(* IEC 61131-3 sources: volt/packages/volt-lsp-iec/test-corpus/lenze-mid/Device/Plc Logic/Application/Library Manager/CAA RTCLK, 21 files *)

(* ---- ERROR.dut ---- *)
TYPE ERROR :
(
	NO_ERROR := 0,
	FIRST_ERROR := 5700,
	TIME_OUT := 5701,
	NOT_AVAILABLE := 5702,
	TIME_NOT_VALID := 5703,
	WRONG_PARAMETER := 5704,
	ERROR_UNKNOWN := 5705,
	NOT_IMPLEMENTED := 5706,
	FIRST_MF := 5725,
	LAST_ERROR := 5749
);
END_TYPE

(* ---- PERIODE.dut ---- *)
TYPE PERIODE :
(
	UNKNOWN := 0,
	STANDARD := 1,
	DAYLIGHT := 2
);
END_TYPE

(* ---- PERIODE_INFO.dut ---- *)
TYPE PERIODE_INFO : RTCLK_PERIODE_INFO;
END_TYPE

(* ---- RTCLK_GETDATEANDTIME_PARAMS.dut ---- *)
TYPE RTCLK_GETDATEANDTIME_PARAMS :
STRUCT
	DTDATEANDTIME : DATE_AND_TIME;
	ETIMEZONE : PERIODE;
END_STRUCT
END_TYPE

(* ---- RTCLK_GETTIMEZONEINFORMATION_PARAMS.dut ---- *)
TYPE RTCLK_GETTIMEZONEINFORMATION_PARAMS :
STRUCT
	TZITIMEZONE : RTCLK_TIME_ZONE_INFO;
END_STRUCT
END_TYPE

(* ---- RTCLK_PERIODE_INFO.dut ---- *)
TYPE RTCLK_PERIODE_INFO :
STRUCT
	SNAME : STRING(32);
	TMDATE : RTCLK_SYSTEMTIME;
	IBIAS : INT;
END_STRUCT
END_TYPE

(* ---- RTCLK_SETDATEANDTIME_PARAMS.dut ---- *)
TYPE RTCLK_SETDATEANDTIME_PARAMS :
STRUCT
	DTDATEANDTIME : DATE_AND_TIME;
END_STRUCT
END_TYPE

(* ---- RTCLK_SETTIMEZONEINFORMATION_PARAMS.dut ---- *)
TYPE RTCLK_SETTIMEZONEINFORMATION_PARAMS :
STRUCT
	TZITIMEZONE : RTCLK_TIME_ZONE_INFO;
END_STRUCT
END_TYPE

(* ---- RTCLK_SYSTEMTIME.dut ---- *)
TYPE RTCLK_SYSTEMTIME :
STRUCT
	UIYEAR : UINT;
	UIMONTH : UINT;
	EWEEKDAY : WEEKDAY;
	UIDAY : UINT;
	UIHOUR : UINT;
	UIMINUTE : UINT;
	UISECOND : UINT;
END_STRUCT
END_TYPE

(* ---- RTCLK_TIME_ZONE_INFO.dut ---- *)
TYPE RTCLK_TIME_ZONE_INFO :
STRUCT
	IBIAS : INT;
	SPERIODE : ARRAY [1..2] OF RTCLK_PERIODE_INFO;
END_STRUCT
END_TYPE

(* ---- SYSTEMTIME.dut ---- *)
TYPE SYSTEMTIME : RTCLK_SYSTEMTIME;
END_TYPE

(* ---- TIME_ZONE_INFO.dut ---- *)
TYPE TIME_ZONE_INFO : RTCLK_TIME_ZONE_INFO;
END_TYPE

(* ---- WEEKDAY.dut ---- *)
TYPE WEEKDAY :
(
	SUNDAY := 0,
	MONDAY := 1,
	TUESDAY := 2,
	WEDNESDAY := 3,
	THURSDAY := 4,
	FRIDAY := 5,
	SATURDAY := 6
);
END_TYPE

(* ---- PROPERTYCONSTANTS.gvl ---- *)
VAR_GLOBAL
	GC_WTIMEZONESUPPORT : WORD := 1;
END_VAR

(* ---- VERSIONCONSTANTS.gvl ---- *)
VAR_GLOBAL
	GC_BYVERSION : BYTE := 1;
	GC_BYVERSION_1 : BYTE := 0;
END_VAR

(* ---- GETPROPERTY.pou ---- *)
FUNCTION GETPROPERTY : __XWORD
VAR_INPUT
	WPROPERTY : WORD;
END_VAR
END_FUNCTION

(* ---- GETSUPPLIERVERSION.pou ---- *)
FUNCTION GETSUPPLIERVERSION : WORD
VAR_INPUT
	XDUMMY : BOOL;
END_VAR
END_FUNCTION

(* ---- GETDATEANDTIME.pou ---- *)
FUNCTION_BLOCK GETDATEANDTIME
VAR_INPUT
	XEXECUTE : BOOL;
END_VAR
VAR_OUTPUT
	XDONE : BOOL;
	XBUSY : BOOL;
	XERROR : BOOL;
	EERROR : ERROR;
	DTDATEANDTIME : DATE_AND_TIME;
	ETIMEZONE : PERIODE;
END_VAR
VAR
	XPREVIOUSEXECUTE : BOOL;
	XPREVIOUSABORTINPROGRESS : BOOL;
	XABORTINPROGRESS : BOOL;
	IERROR : INT;
	HJOB : CAA.HANDLE;
	PGETDATEANDTIMEPARAMS : POINTER TO RTCLK_GETDATEANDTIME_PARAMS;
	STATEJOB : ASM.STATE;
	DWETRIGCLASS : __XWORD;
END_VAR
END_FUNCTION_BLOCK

METHOD FB_EXIT : BOOL
VAR_INPUT
	BINCOPYCODE : BOOL;
END_VAR
END_METHOD

METHOD FB_INIT : BOOL
VAR_INPUT
	BINITRETAINS : BOOL;
	BINCOPYCODE : BOOL;
END_VAR
END_METHOD

(* ---- GETTIMEZONEINFORMATION.pou ---- *)
FUNCTION_BLOCK GETTIMEZONEINFORMATION
VAR_INPUT
	XEXECUTE : BOOL;
END_VAR
VAR_OUTPUT
	XDONE : BOOL;
	XBUSY : BOOL;
	XERROR : BOOL;
	EERROR : ERROR;
	TZIINFO : RTCLK_TIME_ZONE_INFO;
END_VAR
VAR
	XPREVIOUSEXECUTE : BOOL;
	XPREVIOUSABORTINPROGRESS : BOOL;
	XABORTINPROGRESS : BOOL;
	IERROR : INT;
	HJOB : CAA.HANDLE;
	PGETTIMEZONEINFORMATIONPARAMS : POINTER TO RTCLK_GETTIMEZONEINFORMATION_PARAMS;
	STATEJOB : ASM.STATE;
	DWETRIGCLASS : __XWORD;
END_VAR
END_FUNCTION_BLOCK

METHOD FB_EXIT : BOOL
VAR_INPUT
	BINCOPYCODE : BOOL;
END_VAR
END_METHOD

METHOD FB_INIT : BOOL
VAR_INPUT
	BINITRETAINS : BOOL;
	BINCOPYCODE : BOOL;
END_VAR
END_METHOD

(* ---- SETDATEANDTIME.pou ---- *)
FUNCTION_BLOCK SETDATEANDTIME
VAR_INPUT
	XEXECUTE : BOOL;
	DTDATEANDTIME : DATE_AND_TIME;
END_VAR
VAR_OUTPUT
	XDONE : BOOL;
	XBUSY : BOOL;
	XERROR : BOOL;
	EERROR : ERROR;
END_VAR
VAR
	XPREVIOUSEXECUTE : BOOL;
	XPREVIOUSABORTINPROGRESS : BOOL;
	XABORTINPROGRESS : BOOL;
	IERROR : INT;
	HJOB : CAA.HANDLE;
	PSETDATEANDTIMEPARAMS : POINTER TO RTCLK_SETDATEANDTIME_PARAMS;
	STATEJOB : ASM.STATE;
	DWETRIGCLASS : __XWORD;
END_VAR
END_FUNCTION_BLOCK

METHOD FB_EXIT : BOOL
VAR_INPUT
	BINCOPYCODE : BOOL;
END_VAR
END_METHOD

METHOD FB_INIT : BOOL
VAR_INPUT
	BINITRETAINS : BOOL;
	BINCOPYCODE : BOOL;
END_VAR
END_METHOD

(* ---- SETTIMEZONEINFORMATION.pou ---- *)
FUNCTION_BLOCK SETTIMEZONEINFORMATION
VAR_INPUT
	XEXECUTE : BOOL;
	TZIINFO : RTCLK_TIME_ZONE_INFO;
END_VAR
VAR_OUTPUT
	XDONE : BOOL;
	XBUSY : BOOL;
	XERROR : BOOL;
	EERROR : ERROR;
END_VAR
VAR
	XPREVIOUSEXECUTE : BOOL;
	XPREVIOUSABORTINPROGRESS : BOOL;
	XABORTINPROGRESS : BOOL;
	IERROR : INT;
	HJOB : CAA.HANDLE;
	PSETTIMEZONEINFORMATIONPARAMS : POINTER TO RTCLK_SETTIMEZONEINFORMATION_PARAMS;
	STATEJOB : ASM.STATE;
	DWETRIGCLASS : __XWORD;
END_VAR
END_FUNCTION_BLOCK

METHOD FB_EXIT : BOOL
VAR_INPUT
	BINCOPYCODE : BOOL;
END_VAR
END_METHOD

METHOD FB_INIT : BOOL
VAR_INPUT
	BINITRETAINS : BOOL;
	BINCOPYCODE : BOOL;
END_VAR
END_METHOD
